Fanuc KAREL source: kt00304.KL

-- PROVISIONAL review KL for V1013-1; original PC SHA256 d4d6ec057bccf2d9686390d6f18d0e28a5d14b95828918ab74eb64f2c971d56b
-- Incomplete behavior may be omitted. Consult companion uncertainty JSON. Do not deploy.
PROGRAM KT00304
%NOLOCKGROUP
VAR
  R2 : REAL
  OUT : BOOLEAN
-- UNRESOLVED_DECL Y1 type=002018
BEGIN
  -- UNRESOLVED_PC offsets 5-19; opcodes 2E,22,9D,33,B2
  -- UNRESOLVED_PC offsets 24-35; opcodes 2E,23
  -- UNRESOLVED_PC offsets 40-64; opcodes 22,9D,33,B1,21,29,64,6E,23
  -- UNRESOLVED_PC offsets 69-73; opcodes 7F
END KT00304
